(* IEC 61131-3 sources: llm-plc-st-eval/data/raw/gpt-4o/B5/zero_shot, 3 files *)

(* ---- ejec_1.st ---- *)
```pascal
FUNCTION_BLOCK FB_Ventilador
VAR
    // Variable de entrada: estado del quemador
    quemadorOn : BOOL;

    // Variable de salida: estado del ventilador
    ventilador : BOOL;

    // Temporizador para controlar el tiempo de funcionamiento adicional del ventilador
    timer : TON;

    // Variable interna para almacenar el estado previo del quemador
    quemadorPrev : BOOL;
END_VAR

// Inicialización del temporizador
timer(IN := FALSE, PT := T#30S);

// Lógica del ventilador
IF quemadorOn THEN
    // Si el quemador está encendido, el ventilador debe estar encendido
    ventilador := TRUE;
    // Reiniciar el temporizador si el quemador está encendido
    timer(IN := FALSE);
ELSE
    // Si el quemador se apaga, iniciar el temporizador
    IF NOT quemadorPrev THEN
        timer(IN := TRUE);
    END_IF;

    // El ventilador sigue encendido mientras el temporizador está activo
    ventilador := timer.Q;
END_IF;

// Actualizar el estado previo del quemador
quemadorPrev := quemadorOn;
END_FUNCTION_BLOCK
```

Este código implementa la lógica requerida para controlar el ventilador de enfriamiento de un horno. El ventilador se mantiene encendido mientras el quemador está activo y continúa funcionando durante 30 segundos adicionales después de que el quemador se apaga.

(* ---- ejec_2.st ---- *)
```pascal
FUNCTION_BLOCK FB_Ventilador
VAR
    // Variable de entrada: indica si el quemador está encendido
    quemadorOn : BOOL;

    // Variable de salida: controla el estado del ventilador
    ventilador : BOOL;

    // Temporizador para controlar el tiempo adicional de funcionamiento del ventilador
    timer : TON;

    // Variable interna para almacenar el estado anterior del quemador
    quemadorPrev : BOOL;
END_VAR

// Inicialización del temporizador
timer(IN := FALSE, PT := T#30S);

// Lógica de control del ventilador
IF quemadorOn THEN
    // Si el quemador está encendido, el ventilador debe estar encendido
    ventilador := TRUE;
    // Reiniciar el temporizador si el quemador está encendido
    timer(IN := FALSE);
ELSE
    // Si el quemador se apaga, iniciar el temporizador
    IF NOT quemadorPrev THEN
        timer(IN := TRUE);
    END_IF;

    // El ventilador sigue encendido mientras el temporizador no haya alcanzado el tiempo preestablecido
    ventilador := NOT timer.Q;
END_IF;

// Actualizar el estado anterior del quemador
quemadorPrev := quemadorOn;
END_FUNCTION_BLOCK
```

(* ---- ejec_3.st ---- *)
```pascal
FUNCTION_BLOCK FB_Ventilador
VAR
    // Variable de entrada
    quemadorOn : BOOL; // Estado del quemador: TRUE si está encendido, FALSE si está apagado

    // Variable de salida
    ventilador : BOOL; // Estado del ventilador: TRUE si está encendido, FALSE si está apagado

    // Variables internas
    timer : TON; // Temporizador para controlar el tiempo adicional de funcionamiento del ventilador
END_VAR

// Inicialización del temporizador
timer(IN := NOT quemadorOn, PT := T#30S);

// Lógica de control del ventilador
IF quemadorOn THEN
    ventilador := TRUE; // El ventilador está encendido mientras el quemador está encendido
ELSE
    timer(IN := TRUE); // Iniciar el temporizador cuando el quemador se apaga
    ventilador := timer.Q; // El ventilador sigue encendido mientras el temporizador está activo
END_IF;
```

Este código define un bloque de función `FB_Ventilador` que controla el estado de un ventilador de enfriamiento basado en el estado de un quemador. Utiliza un temporizador `TON` para mantener el ventilador encendido durante 30 segundos después de que el quemador se apague.
